(* IEC 61131-3 sources: Gen-AI/release/member2-v1.1/成员2_提交包_v1.1/agent/logs/scenario_fixture/timeout/fixture/E3_S03_1_42, 3 files *)

(* ---- best.st ---- *)
FUNCTION_BLOCK FB_S03
VAR_INPUT
    DoorSwitch : BOOL;
    ZoneAOccupied : BOOL;
    ZoneBOccupied : BOOL;
    ResetBtn : BOOL;
    EStop_NC : BOOL;
END_VAR
VAR_OUTPUT
    DriveA_Run : BOOL;
    DriveB_Run : BOOL;
    AlarmLamp : BOOL;
    Status : WORD;
END_VAR
(* Add a VAR block for internal state/timers before the implementation, if needed. *)
(* SKELETON ONLY: replace this RETURN with scan logic and required initial state. *)
RETURN;
END_FUNCTION_BLOCK

(* FIXTURE_TIMEOUT *)

(* ---- final.st ---- *)
FUNCTION_BLOCK FB_S03
VAR_INPUT
    DoorSwitch : BOOL;
    ZoneAOccupied : BOOL;
    ZoneBOccupied : BOOL;
    ResetBtn : BOOL;
    EStop_NC : BOOL;
END_VAR
VAR_OUTPUT
    DriveA_Run : BOOL;
    DriveB_Run : BOOL;
    AlarmLamp : BOOL;
    Status : WORD;
END_VAR
(* Add a VAR block for internal state/timers before the implementation, if needed. *)
(* SKELETON ONLY: replace this RETURN with scan logic and required initial state. *)
RETURN;
END_FUNCTION_BLOCK

(* FIXTURE_TIMEOUT *)

(* ---- skeleton.st ---- *)
FUNCTION_BLOCK FB_S03
VAR_INPUT
    DoorSwitch : BOOL;
    ZoneAOccupied : BOOL;
    ZoneBOccupied : BOOL;
    ResetBtn : BOOL;
    EStop_NC : BOOL;
END_VAR
VAR_OUTPUT
    DriveA_Run : BOOL;
    DriveB_Run : BOOL;
    AlarmLamp : BOOL;
    Status : WORD;
END_VAR
(* Add a VAR block for internal state/timers before the implementation, if needed. *)
(* SKELETON ONLY: replace this RETURN with scan logic and required initial state. *)
RETURN;
END_FUNCTION_BLOCK
